(* IEC 61131-3 sources: BODAS-HelloWorld/st/bodas_rc18_12_40/plc_logic/application/01_maintask/11_parameters/programs, 1 file *)

(* ---- prg_nvmconfig-PRG_NVMConfig.st ---- *)
(* --- Interface --- *)
(*********************************************************************************************************************
 *     __   __   ___  ___           __   __        __   __  ___
 *   /_ / /  / /__  /    /__/     /_ / /_   |_ / /_ / /  /  /  /__/
 *  /__/ /__/ __ / /__  /  /     /  | /__  /  | /  | /__/  /  /  /
 *
 * Project: Hello World for ml290.rts
 *
 * Program: PRG_NVMConfig
 *
 * Author:
 *
 * Description:
 * Interface for Paramters
 *
 * (c) Copyright by BOSCH REXROTH AG, all rights reserved
 *
 *********************************************************************************************************************)
PROGRAM PRG_NVMConfig
VAR
	status_u16 : UINT;
END_VAR

(* --- Implementation --- *)
;
